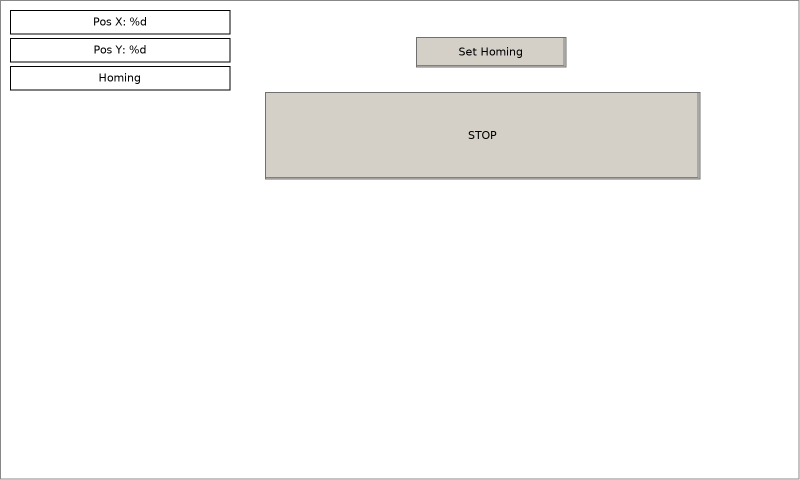
VISUALIZATION VisuTest  // 800x480
    Rectangle (10,10 220x24), "Pos X: %d", text variable: MAIN.CurrentPosX
    Rectangle (10,38 220x24), "Pos Y: %d", text variable: MAIN.CurrentPosY
    Rectangle (10,66 220x24), "Homing", colour toggle: MAIN.isHoming
    Button (416,37 150x30), "Set Homing"
        OnMouseDown: toggle MAIN.isHoming
    Button (265,92 435x87), "STOP"
        OnMouseDown: execute {
            Main.M2_Forward := FALSE;
            Main.M2_Back    := FALSE;
            Main.M3_Down    := FALSE;
            Main.M3_Up      := FALSE;
            Main.M4_Forward := FALSE;
            Main.M4_Back    := FALSE;
        }
END_VISUALIZATION

(* stored: Version 1.1.0.1, ProductVersion 3.1.4024.12
   Visu VisuTest: Id {6e3f99c2-464f-4e1a-aa55-836022e67384} *)
